// TIA Portal V21 export
// export: Created 2026-11-22T00:27:48.0708534Z, ExportSetting WithDefaults, DisplayName Totally Integrated Automation Portal, DisplayVersion V21 Update 3, DisplayName STEP 7 Professional, DisplayVersion V21 Update 3, DisplayName STEP 7 Safety, DisplayVersion V21, DisplayName Tech WebApplication, DisplayVersion V21, DisplayName WinCC Basic/Comfort/Advanced, DisplayVersion V21 Update 3, DisplayName WinCC Unified, DisplayVersion V21 Update 3
Screen "P_Clock_2"  1280x800, Number=120
  ScreenLayer "Layer_0"
    Clock "TicksColor" at 10,10 size 150x150  TickDistance=80, StyleItem=Clock
    TextField "Label_TicksColor" at 10,162 size 158x16  StyleItem=Text field, Text="TicksColor"
    Clock "UseDesignColorSchema" at 170,10 size 150x150  TickDistance=80
    TextField "Label_UseDesignColorSchema" at 170,162 size 158x16  StyleItem=Text field, Text="UseDesignColorSchema"
    Button "Next" at 1238,776 size 40x22  Mode=Text, StyleItem=Button, TextOff="Text", TextOn="Text"
      on Click: ActivateScreen(Screen name := P_Line_1, Object number := 0)
